# EPICS substitutions: db/Beckhoff_5XXX/ecmcEL5001.substitutions
file "ecmcEL500X-chX.template"
{
  pattern {CH_ID}
          {01   }
}
